PROGRAM Init
VAR
	bFirstTime					:BOOL; 				(* False = first run / True = not first run *)
END_VAR
VAR PERSISTENT
	bFirstTimePersistent			:BOOL;				(* Persistente Daten initialisieren *)
END_VAR


IF NOT bFirstTime
THEN
	A_InitGr0000();
	A_InitGr0100();
	A_InitGr0200();
	A_InitGr0500();

	bFirstTime:= TRUE;
END_IF

IF NOT bFirstTimePersistent
THEN

	bFirstTimePersistent:= TRUE;
END_IF

ACTION A_InitGr0000:
;
END_ACTION

ACTION A_InitGr0100:
;
END_ACTION

ACTION A_InitGr0200:
;
END_ACTION

ACTION A_InitGr0500:
;
END_ACTION

END_PROGRAM

(* stored: Version 1.1.0.1, ProductVersion 3.1.4024.15
   POU Init: Id {686a804b-e730-4808-9911-31ba1cd60631}, SpecialFunc None
   Action A_InitGr0000: Id {63a26e6c-4076-4d09-8cff-2202182e2987}
   Action A_InitGr0100: Id {2c5d6dff-d3bb-4929-83d0-4de6332805af}
   Action A_InitGr0200: Id {2e59a8af-7993-4673-973b-1fa912614abb}
   Action A_InitGr0500: Id {962e3661-f1b0-4ae8-aef7-cf49232dcb82} *)
